Fanuc KAREL source: NC0084.KL

PROGRAM NC0084
%NOLOCKGROUP
ROUTINE R
VAR
S1:INTEGER;S2:INTEGER
BEGIN
--
S1=1
IF (S1=1) THEN
SELECT S1 OF
CASE(1):
FOR S2=1 TO 2 DO
S1=(S1+1)
ENDFOR
CASE(2):
S1=(S1+2)
ELSE:
S1=(S1+3)
ENDSELECT
ELSE
S1=(S1+2)
ENDIF
END R
BEGIN
R
END NC0084
